Fanuc KAREL source: kb00176.compact.KL

PROGRAM KB00176
%STACKSIZE=65535
%PRIORITY=65535
%NOLOCKGROUP
%ENVIRONMENT REGOPE
VAR
P1 : INTEGER
P2 : XYZWPR
P3 : INTEGER
BEGIN
P1=1
P2.X=1.0
P3=1
SET_POS_REG(P1,P2,P3,1)
END KB00176
